(* IEC 61131-3 sources: ConveyorControl-with-PLC/4E_Gruppe1_Graf_Projekt1/Drive, 3 files *)

(* ---- _DriveAxis1.st ---- *)
FUNCTION GLOBAL TAB DRIVETAB__DRIVEAXIS1_0
	1$UDINT, TO_UDINT(OFF(L1)-OFF(L0)),L0:
G01:	1$USINT,' '' '' '' ',
	2$USINT,' '' '' '' ',
	3$USINT,' '' '' '' ',
	4$USINT,460$DINT,
	5$USINT,920$DINT,
	6$USINT,2750$DINT,
	7$USINT,6$DINT,
	8$USINT,1700$DINT,
	9$USINT,1000$DINT,
	10$USINT,1000$DINT,
	11$USINT,10$DINT,
	12$USINT,517$DINT,
	13$USINT,2$DINT,
	14$USINT,0$DINT,
	15$USINT,1024$DINT,
	16$USINT,1500$DINT,
	17$USINT,0$DINT,
	18$USINT,0$DINT,
	21$USINT,0$DINT,
	22$USINT,10$DINT,
	23$USINT,10$DINT,
	24$USINT,230$DINT,
	25$USINT,11$DINT,
	26$USINT,0$DINT,
	27$USINT,20$DINT,
G03:	32$USINT,2$DINT,
	33$USINT,50$DINT,
	34$USINT,480$DINT,
	35$USINT,100$DINT,
	36$USINT,200$DINT,
	37$USINT,85$DINT,
	38$USINT,85$DINT,
	39$USINT,1$DINT,
	40$USINT,1$DINT,
	41$USINT,65$DINT,
	42$USINT,2750$DINT,
	43$USINT,2621740$DINT,
	44$USINT,966188242$DINT,
	45$USINT,-1035927552$DINT,
	46$USINT,67117569$DINT,
	47$USINT,2750$DINT,
	48$USINT,1$DINT,
	49$USINT,25$DINT,
	168$USINT,60$DINT,
	169$USINT,55$DINT,
	170$USINT,55$DINT,
G04:	50$USINT,100000$DINT,
	51$USINT,1000$DINT,
	52$USINT,30$DINT,
	53$USINT,70$DINT,
	54$USINT,70$DINT,
	55$USINT,40$DINT,
	56$USINT,460$DINT,
	57$USINT,920$DINT,
	58$USINT,920$DINT,
G05:	60$USINT,5000$DINT,
	61$USINT,10000$DINT,
	62$USINT,400$DINT,
	63$USINT,1000$DINT,
	64$USINT,80$DINT,
	65$USINT,2750$DINT,
	66$USINT,0$DINT,
G06:	70$USINT,20000$DINT,
	71$USINT,1000$DINT,
	72$USINT,0$DINT,
	73$USINT,1000$DINT,
	74$USINT,0$DINT,
	75$USINT,2147483647$DINT,
	76$USINT,0$DINT,
G07:	80$USINT,600$DINT,
	81$USINT,0$DINT,
	82$USINT,0$DINT,
G08:	90$USINT,1000$DINT,
	91$USINT,517$DINT,
	92$USINT,0$DINT,
	93$USINT,2562$DINT,
	94$USINT,0$DINT,
	95$USINT,1000$DINT,
	96$USINT,250$DINT,
	97$USINT,0$DINT,
	98$USINT,0$DINT,
	99$USINT,100$DINT,
	100$USINT,0$DINT,
	101$USINT,100$DINT,
	102$USINT,0$DINT,
	103$USINT,0$DINT,
	104$USINT,0$DINT,
	105$USINT,0$DINT,
	106$USINT,0$DINT,
	107$USINT,0$DINT,
	108$USINT,' '' '' '' ',
	109$USINT,' '' '' '' ',
	110$USINT,' '' '' '' ',
	111$USINT,0$DINT,
	112$USINT,0$DINT,
	113$USINT,0$DINT,
	114$USINT,0$DINT,
	115$USINT,0$DINT,
	116$USINT,0$DINT,
	117$USINT,100$DINT,
	118$USINT,0$DINT,
	119$USINT,2500$DINT,
	120$USINT,300$DINT,
	121$USINT,2000$DINT,
	122$USINT,0$DINT,L1:
TO_UDINT(OFF(L3)-OFF(L2)),L2:
	01$USINT, OFF(G01),
	03$USINT, OFF(G03),
	04$USINT, OFF(G04),
	05$USINT, OFF(G05),
	06$USINT, OFF(G06),
	07$USINT, OFF(G07),
	08$USINT, OFF(G08),L3:
END_FUNCTION

(* ---- _DriveAxis1_01.st ---- *)
FUNCTION GLOBAL TAB DRIVETAB__DRIVEAXIS1_1
	1$UDINT, TO_UDINT(OFF(L1)-OFF(L0)),L0:
G01:	1$USINT,' '' '' '' ',
	2$USINT,' '' '' '' ',
	3$USINT,' '' '' '' ',
	4$USINT,460$DINT,
	5$USINT,920$DINT,
	6$USINT,2750$DINT,
	7$USINT,6$DINT,
	8$USINT,1700$DINT,
	9$USINT,1000$DINT,
	10$USINT,1000$DINT,
	11$USINT,10$DINT,
	12$USINT,517$DINT,
	13$USINT,2$DINT,
	14$USINT,0$DINT,
	15$USINT,1024$DINT,
	16$USINT,1500$DINT,
	17$USINT,0$DINT,
	18$USINT,0$DINT,
	21$USINT,0$DINT,
	22$USINT,10$DINT,
	23$USINT,10$DINT,
	24$USINT,230$DINT,
	25$USINT,11$DINT,
	26$USINT,0$DINT,
	27$USINT,20$DINT,
G03:	32$USINT,2$DINT,
	33$USINT,50$DINT,
	34$USINT,230$DINT,
	35$USINT,100$DINT,
	36$USINT,33$DINT,
	37$USINT,85$DINT,
	38$USINT,85$DINT,
	39$USINT,1$DINT,
	40$USINT,1$DINT,
	41$USINT,65$DINT,
	42$USINT,2750$DINT,
	43$USINT,2621740$DINT,
	44$USINT,966188242$DINT,
	45$USINT,-1035927552$DINT,
	46$USINT,67117569$DINT,
	47$USINT,2750$DINT,
	48$USINT,1$DINT,
	49$USINT,100$DINT,
	168$USINT,60$DINT,
	169$USINT,55$DINT,
	170$USINT,55$DINT,
G04:	50$USINT,100000$DINT,
	51$USINT,1000$DINT,
	52$USINT,30$DINT,
	53$USINT,70$DINT,
	54$USINT,70$DINT,
	55$USINT,40$DINT,
	56$USINT,460$DINT,
	57$USINT,920$DINT,
	58$USINT,920$DINT,
G05:	60$USINT,5000$DINT,
	61$USINT,10000$DINT,
	62$USINT,400$DINT,
	63$USINT,1000$DINT,
	64$USINT,80$DINT,
	65$USINT,2750$DINT,
	66$USINT,0$DINT,
G06:	70$USINT,20000$DINT,
	71$USINT,1000$DINT,
	72$USINT,0$DINT,
	73$USINT,1000$DINT,
	74$USINT,0$DINT,
	75$USINT,2147483647$DINT,
	76$USINT,0$DINT,
G07:	80$USINT,600$DINT,
	81$USINT,0$DINT,
	82$USINT,0$DINT,
G08:	90$USINT,1000$DINT,
	91$USINT,517$DINT,
	92$USINT,0$DINT,
	93$USINT,2562$DINT,
	94$USINT,0$DINT,
	95$USINT,1000$DINT,
	96$USINT,250$DINT,
	97$USINT,0$DINT,
	98$USINT,0$DINT,
	99$USINT,100$DINT,
	100$USINT,0$DINT,
	101$USINT,100$DINT,
	102$USINT,0$DINT,
	103$USINT,0$DINT,
	104$USINT,0$DINT,
	105$USINT,0$DINT,
	106$USINT,0$DINT,
	107$USINT,0$DINT,
	108$USINT,' '' '' '' ',
	109$USINT,' '' '' '' ',
	110$USINT,' '' '' '' ',
	111$USINT,0$DINT,
	112$USINT,0$DINT,
	113$USINT,0$DINT,
	114$USINT,0$DINT,
	115$USINT,0$DINT,
	116$USINT,0$DINT,
	117$USINT,100$DINT,
	118$USINT,0$DINT,
	119$USINT,2500$DINT,
	120$USINT,300$DINT,
	121$USINT,2000$DINT,
	122$USINT,0$DINT,L1:
TO_UDINT(OFF(L3)-OFF(L2)),L2:
	01$USINT, OFF(G01),
	03$USINT, OFF(G03),
	04$USINT, OFF(G04),
	05$USINT, OFF(G05),
	06$USINT, OFF(G06),
	07$USINT, OFF(G07),
	08$USINT, OFF(G08),L3:
END_FUNCTION

(* ---- _DriveAxis2.st ---- *)
FUNCTION GLOBAL TAB DRIVETAB__DRIVEAXIS2
	1$UDINT, TO_UDINT(OFF(L1)-OFF(L0)),L0:
G01:	1$USINT,' '' '' '' ',
	2$USINT,' '' '' '' ',
	3$USINT,' '' '' '' ',
	4$USINT,5000$DINT,
	5$USINT,10000$DINT,
	6$USINT,3000$DINT,
	7$USINT,6$DINT,
	8$USINT,1700$DINT,
	9$USINT,1000$DINT,
	10$USINT,1000$DINT,
	11$USINT,10$DINT,
	12$USINT,0$DINT,
	13$USINT,2$DINT,
	14$USINT,0$DINT,
	15$USINT,1024$DINT,
	16$USINT,1500$DINT,
	17$USINT,0$DINT,
	18$USINT,0$DINT,
	21$USINT,0$DINT,
	22$USINT,10$DINT,
	23$USINT,100$DINT,
	24$USINT,0$DINT,
	25$USINT,0$DINT,
	26$USINT,0$DINT,
	27$USINT,20$DINT,
G03:	32$USINT,3$DINT,
	33$USINT,50$DINT,
	34$USINT,480$DINT,
	35$USINT,100$DINT,
	36$USINT,200$DINT,
	37$USINT,85$DINT,
	38$USINT,85$DINT,
	39$USINT,0$DINT,
	40$USINT,0$DINT,
	41$USINT,65$DINT,
	42$USINT,10000$DINT,
	43$USINT,2621740$DINT,
	44$USINT,999808723$DINT,
	45$USINT,1077936128$DINT,
	46$USINT,67117056$DINT,
	47$USINT,300000$DINT,
	48$USINT,1$DINT,
	49$USINT,25$DINT,
	168$USINT,60$DINT,
	169$USINT,55$DINT,
	170$USINT,55$DINT,
G04:	50$USINT,25000$DINT,
	51$USINT,1000$DINT,
	52$USINT,30$DINT,
	53$USINT,70$DINT,
	54$USINT,70$DINT,
	55$USINT,40$DINT,
	56$USINT,0$DINT,
	57$USINT,0$DINT,
	58$USINT,0$DINT,
G05:	60$USINT,5000$DINT,
	61$USINT,10000$DINT,
	62$USINT,400$DINT,
	63$USINT,1000$DINT,
	64$USINT,80$DINT,
	65$USINT,3000$DINT,
	66$USINT,0$DINT,
G06:	70$USINT,20000$DINT,
	71$USINT,1000$DINT,
	72$USINT,16$DINT,
	73$USINT,1000$DINT,
	74$USINT,0$DINT,
	75$USINT,327680$DINT,
	76$USINT,0$DINT,
G07:	80$USINT,600$DINT,
	81$USINT,0$DINT,
	82$USINT,0$DINT,
G08:	90$USINT,5000$DINT,
	91$USINT,775$DINT,
	92$USINT,0$DINT,
	93$USINT,3591$DINT,
	94$USINT,0$DINT,
	95$USINT,4000$DINT,
	96$USINT,250$DINT,
	97$USINT,0$DINT,
	98$USINT,0$DINT,
	99$USINT,100$DINT,
	100$USINT,0$DINT,
	101$USINT,100$DINT,
	102$USINT,75$DINT,
	103$USINT,100$DINT,
	104$USINT,0$DINT,
	105$USINT,0$DINT,
	106$USINT,0$DINT,
	107$USINT,0$DINT,
	108$USINT,' '' '' '' ',
	109$USINT,' '' '' '' ',
	110$USINT,' '' '' '' ',
	111$USINT,0$DINT,
	112$USINT,0$DINT,
	113$USINT,0$DINT,
	114$USINT,0$DINT,
	115$USINT,0$DINT,
	116$USINT,0$DINT,
	117$USINT,100$DINT,
	118$USINT,0$DINT,
	119$USINT,2500$DINT,
	120$USINT,300$DINT,
	121$USINT,2000$DINT,
	122$USINT,0$DINT,L1:
TO_UDINT(OFF(L3)-OFF(L2)),L2:
	01$USINT, OFF(G01),
	03$USINT, OFF(G03),
	04$USINT, OFF(G04),
	05$USINT, OFF(G05),
	06$USINT, OFF(G06),
	07$USINT, OFF(G07),
	08$USINT, OFF(G08),L3:
END_FUNCTION
